// TIA Portal V21 export
DATA_BLOCK "Issue221_root_omitted"   // DB
// stored: AutoNumber true
BEGIN
END_DATA_BLOCK
